Staubli VAL3: login.pgx

public program login(bool& x_bResult)
  local bool l_bCancel
begin
  sPage=""
  x_bResult=false
  do
    if sPage!="login"
      sPage="login"
      //init
      sInputPswd=""
      //bind
      userPageBind("login","pwd1","value",sInputPswd,1,"rw")
      userPageBindClick("login","btn1",bConfirm,true)
      userPageBindClick("login","btn2",bCancel,true)
      //
      userPage(sPage)
      delay(0.5)
    endIf
    //button
    if bConfirm
      bConfirm=false
      if sInputPswd==sPassword
        x_bResult=true
      else
        userPageAlert("invalid password!")
      endIf
    elseIf bCancel
      bCancel=false
      l_bCancel=true
    endIf




    delay(0)
  until l_bCancel==true
end
